Staubli VAL3: checkPoint.pgx

public program checkPoint()
  local num l_nSize
  local num l_i
  local pointRx l_pPoint
  local bool l_bErr
begin
  l_pPoint=here(flange,world)
  l_nSize=size(safeData:sSPoint)
  for l_i = 0 to l_nSize-1
    if safeData:sSPoint[l_i].bActive
      if distance(safeData:sSPoint[l_i].pPointRx.trsf,l_pPoint.trsf)<5
        call io:setDigOutput(io:dOutput[l_i+96],true,l_bErr)
      else
        call io:setDigOutput(io:dOutput[l_i+96],false,l_bErr)
      endIf
    endIf
  endFor
end
